Fanuc KAREL source: kb00039.KL

PROGRAM KB00039
%STACKSIZE=65535
%PRIORITY=65535
%NOLOCKGROUP
VAR
P1 : STRING[80]
P3 : INTEGER
-- UNRESOLVED DECLARATIONS (source type spelling not recovered)
-- P2 : TYPE_0x001C (type_u16=0x001C)
BEGIN
P1='A'
P3=1
CNV_STR_CONF(P1,P2,P3)
END KB00039
